FUNCTION_BLOCK BeltMaster (* Basic Function Block Type *)
  (* Standard: 61499-2 *)
  (* Version 0.0, 11/22/2026, Schneider Electric, First version *)
  PACKAGE Main;
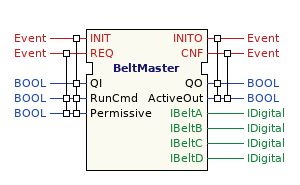
  EVENT_INPUT
    INIT WITH QI, RunCmd, Permissive; (* Initialization Request *)
    REQ WITH RunCmd, Permissive; (* Update belt master setpoint *)
  END_EVENT
  EVENT_OUTPUT
    INITO WITH QO, ActiveOut; (* Initialization Confirm *)
    CNF WITH ActiveOut; (* Execution Confirmation *)
  END_EVENT
  VAR_INPUT
    QI : BOOL := TRUE; (* Input event qualifier *)
    RunCmd : BOOL := FALSE; (* Master belt run command from HMI SetBool *)
    Permissive : BOOL := TRUE; (* Master belt permissive *)
  END_VAR
  VAR_OUTPUT
    QO : BOOL; (* Output event qualifier *)
    ActiveOut : BOOL; (* Effective belt run command *)
  END_VAR
  PLUGS
    IBeltA : IDigital; (* Remote setpoint adapter for BeltA *)
    IBeltB : IDigital; (* Remote setpoint adapter for BeltB *)
    IBeltC : IDigital; (* Remote setpoint adapter for BeltC *)
    IBeltD : IDigital; (* Remote setpoint adapter for BeltD *)
  END_PLUGS
  VAR
    firstFbDoneA : BOOL := FALSE; (* Initial REQ_FB sync completed for BeltA *)
    firstFbDoneB : BOOL := FALSE; (* Initial REQ_FB sync completed for BeltB *)
    firstFbDoneC : BOOL := FALSE; (* Initial REQ_FB sync completed for BeltC *)
    firstFbDoneD : BOOL := FALSE; (* Initial REQ_FB sync completed for BeltD *)
    prevTrackA : BOOL := FALSE; (* Previous Track state for BeltA *)
    prevTrackB : BOOL := FALSE; (* Previous Track state for BeltB *)
    prevTrackC : BOOL := FALSE; (* Previous Track state for BeltC *)
    prevTrackD : BOOL := FALSE; (* Previous Track state for BeltD *)
    targetInt : INT := 0; (* Target integer setpoint (0=Stop, 1=Run) *)
  END_VAR
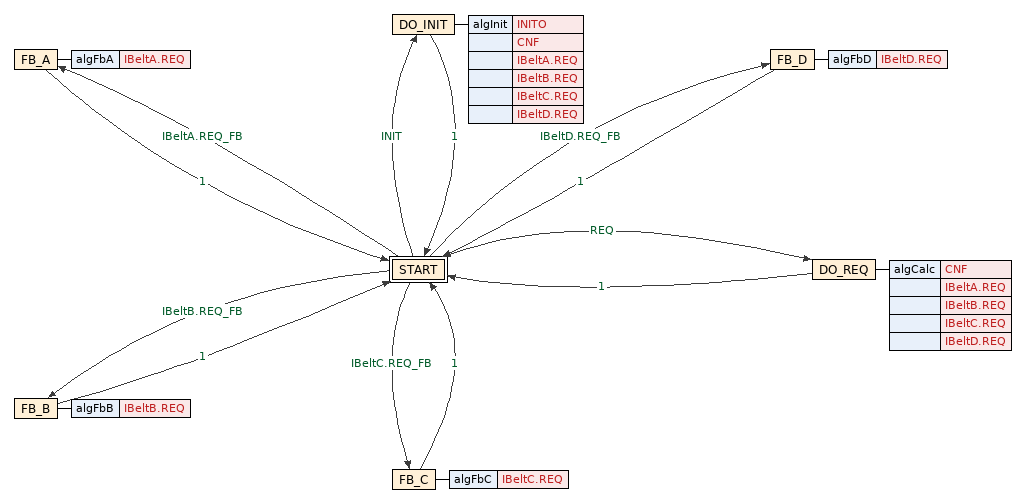
  EC_STATES
    START; (* Initial State *)
    DO_INIT : algInit -> INITO, -> CNF, -> IBeltA.REQ, -> IBeltB.REQ, -> IBeltC.REQ, -> IBeltD.REQ;
    DO_REQ : algCalc -> CNF, -> IBeltA.REQ, -> IBeltB.REQ, -> IBeltC.REQ, -> IBeltD.REQ;
    FB_A : algFbA -> IBeltA.REQ;
    FB_B : algFbB -> IBeltB.REQ;
    FB_C : algFbC -> IBeltC.REQ;
    FB_D : algFbD -> IBeltD.REQ;
  END_STATES
  EC_TRANSITIONS
    START TO DO_INIT := INIT;
    DO_INIT TO START := 1;
    START TO DO_REQ := REQ;
    DO_REQ TO START := 1;
    START TO FB_A := IBeltA.REQ_FB;
    FB_A TO START := 1;
    START TO FB_B := IBeltB.REQ_FB;
    FB_B TO START := 1;
    START TO FB_C := IBeltC.REQ_FB;
    FB_C TO START := 1;
    START TO FB_D := IBeltD.REQ_FB;
    FB_D TO START := 1;
  END_TRANSITIONS
  ALGORITHM algInit IN ST: (* Initialize outputs and push startup setpoints to all 4 belts *)
QO := QI;
ActiveOut := RunCmd AND Permissive;
IF ActiveOut THEN
	targetInt := 1;
ELSE
	targetInt := 0;
END_IF;

IBeltA.Value.value := targetInt;
IBeltA.Value.quality := 16#0;
IBeltB.Value.value := targetInt;
IBeltB.Value.quality := 16#0;
IBeltC.Value.value := targetInt;
IBeltC.Value.quality := 16#0;
IBeltD.Value.value := targetInt;
IBeltD.Value.quality := 16#0;
  END_ALGORITHM
  ALGORITHM algCalc IN ST: (* Compute master belt command and write all 4 belt plugs *)
ActiveOut := RunCmd AND Permissive;
IF ActiveOut THEN
	targetInt := 1;
ELSE
	targetInt := 0;
END_IF;

IBeltA.Value.value := targetInt;
IBeltA.Value.quality := 16#0;
IBeltB.Value.value := targetInt;
IBeltB.Value.quality := 16#0;
IBeltC.Value.value := targetInt;
IBeltC.Value.quality := 16#0;
IBeltD.Value.value := targetInt;
IBeltD.Value.quality := 16#0;
  END_ALGORITHM
  ALGORITHM algFbA IN ST: (* Sync BeltA remote setpoint on first feedback or return to Program Remote *)
IBeltA.REQ := FALSE;
IF (NOT IBeltA.Track) AND ((NOT firstFbDoneA) OR prevTrackA) THEN
	firstFbDoneA := TRUE;
	IBeltA.Value.value := targetInt;
	IBeltA.Value.quality := 16#0;
	IBeltA.REQ := TRUE;
END_IF;
prevTrackA := IBeltA.Track;
  END_ALGORITHM
  ALGORITHM algFbB IN ST: (* Sync BeltB remote setpoint on first feedback or return to Program Remote *)
IBeltB.REQ := FALSE;
IF (NOT IBeltB.Track) AND ((NOT firstFbDoneB) OR prevTrackB) THEN
	firstFbDoneB := TRUE;
	IBeltB.Value.value := targetInt;
	IBeltB.Value.quality := 16#0;
	IBeltB.REQ := TRUE;
END_IF;
prevTrackB := IBeltB.Track;
  END_ALGORITHM
  ALGORITHM algFbC IN ST: (* Sync BeltC remote setpoint on first feedback or return to Program Remote *)
IBeltC.REQ := FALSE;
IF (NOT IBeltC.Track) AND ((NOT firstFbDoneC) OR prevTrackC) THEN
	firstFbDoneC := TRUE;
	IBeltC.Value.value := targetInt;
	IBeltC.Value.quality := 16#0;
	IBeltC.REQ := TRUE;
END_IF;
prevTrackC := IBeltC.Track;
  END_ALGORITHM
  ALGORITHM algFbD IN ST: (* Sync BeltD remote setpoint on first feedback or return to Program Remote *)
IBeltD.REQ := FALSE;
IF (NOT IBeltD.Track) AND ((NOT firstFbDoneD) OR prevTrackD) THEN
	firstFbDoneD := TRUE;
	IBeltD.Value.value := targetInt;
	IBeltD.Value.quality := 16#0;
	IBeltD.REQ := TRUE;
END_IF;
prevTrackD := IBeltD.Track;
  END_ALGORITHM
END_FUNCTION_BLOCK
